(* IEC 61131-3 sources: llm-plc-st-eval/data/definitivo/claude-sonnet-4-6/B6/few_shot, 3 files *)

(* ---- ejec_1.st ---- *)
```st
FUNCTION_BLOCK FB_Baliza
VAR_INPUT
    alarma : BOOL; (* Condicion de alarma activa *)
END_VAR
VAR_OUTPUT
    lampara : BOOL; (* Lampara de baliza *)
END_VAR
VAR
    tOn  : TON; (* Temporizador fase encendida *)
    tOff : TON; (* Temporizador fase apagada *)
    parpadeo : BOOL; (* Estado interno de parpadeo *)
END_VAR

(* Sin alarma: lampara apagada y temporizadores reiniciados *)
IF NOT alarma THEN
    parpadeo := FALSE;
    tOn(IN := FALSE, PT := T#1S);
    tOff(IN := FALSE, PT := T#1S);
ELSE
    (* Fase encendida: activa tOn mientras parpadeo=TRUE *)
    tOn(IN := parpadeo, PT := T#1S);
    (* Fase apagada: activa tOff cuando tOn ha completado *)
    tOff(IN := tOn.Q, PT := T#1S);

    (* Al completar fase apagada, reinicia tOn para nuevo ciclo *)
    IF tOff.Q THEN
        tOn(IN := FALSE, PT := T#1S);  (* Reinicia tOn *)
        tOff(IN := FALSE, PT := T#1S); (* Reinicia tOff *)
        parpadeo := TRUE;
    END_IF;

    (* Arranca el primer ciclo *)
    IF NOT parpadeo AND NOT tOn.Q AND NOT tOff.Q THEN
        parpadeo := TRUE;
    END_IF;
END_IF;

(* La lampara sigue el estado de parpadeo mientras tOn no haya terminado *)
lampara := alarma AND parpadeo AND NOT tOn.Q;
END_FUNCTION_BLOCK
```

(* ---- ejec_2.st ---- *)
```st
FUNCTION_BLOCK FB_Baliza
VAR_INPUT
    alarma : BOOL; (* Condicion de alarma activa *)
END_VAR
VAR_OUTPUT
    lampara : BOOL; (* Lampara de baliza *)
END_VAR
VAR
    tOn  : TON; (* Temporizador fase encendida *)
    tOff : TON; (* Temporizador fase apagada *)
    parpadeo : BOOL; (* Estado interno de parpadeo *)
END_VAR

(* Sin alarma: lampara apagada y temporizadores reiniciados *)
IF NOT alarma THEN
    parpadeo := FALSE;
    tOn(IN := FALSE, PT := T#1S);
    tOff(IN := FALSE, PT := T#1S);
ELSE
    (* Fase encendida: activa tOn mientras parpadeo=TRUE *)
    tOn(IN := parpadeo, PT := T#1S);

    (* Fase apagada: activa tOff cuando tOn ha completado *)
    tOff(IN := tOn.Q, PT := T#1S);

    (* Al completar tOff, reinicia tOn para el siguiente ciclo *)
    IF tOff.Q THEN
        tOn(IN := FALSE, PT := T#1S);  (* Reinicia tOn *)
        tOff(IN := FALSE, PT := T#1S); (* Reinicia tOff *)
        parpadeo := TRUE;
    END_IF;

    (* Arranca el primer ciclo *)
    IF NOT parpadeo AND NOT tOn.Q AND NOT tOff.Q THEN
        parpadeo := TRUE;
    END_IF;
END_IF;

(* La lampara sigue el estado de parpadeo durante la fase encendida *)
lampara := alarma AND parpadeo AND NOT tOn.Q;
END_FUNCTION_BLOCK
```

(* ---- ejec_3.st ---- *)
```pascal
FUNCTION_BLOCK FB_Baliza
VAR_INPUT
    alarma : BOOL; (* Condicion de alarma activa *)
END_VAR
VAR_OUTPUT
    lampara : BOOL; (* Lampara de baliza *)
END_VAR
VAR
    tOn  : TON; (* Temporizador fase encendida *)
    tOff : TON; (* Temporizador fase apagada *)
    parpadeo : BOOL; (* Estado interno de parpadeo *)
END_VAR

(* Sin alarma: lampara apagada y temporizadores reiniciados *)
IF NOT alarma THEN
    parpadeo := FALSE;
    tOn(IN := FALSE, PT := T#1S);
    tOff(IN := FALSE, PT := T#1S);
ELSE
    (* Fase encendida: activa tOn mientras parpadeo=TRUE *)
    tOn(IN := parpadeo, PT := T#1S);

    (* Fase apagada: activa tOff cuando tOn ha completado *)
    tOff(IN := tOn.Q, PT := T#1S);

    (* Al completar tOff vuelve a fase encendida *)
    IF tOff.Q THEN
        parpadeo := FALSE; (* Reinicia para re-disparar tOn *)
    END_IF;

    (* Inicia ciclo: si ninguno esta corriendo, arranca fase encendida *)
    IF NOT tOn.IN AND NOT tOff.IN THEN
        parpadeo := TRUE;
    END_IF;
END_IF;

(* La lampara sigue el estado de parpadeo interno *)
lampara := parpadeo AND alarma;
END_FUNCTION_BLOCK
```
